FUNCTION_BLOCK LiftBootSync (* Basic Function Block Type *)
  (* Standard: 61499-2 *)
  (* Version 0.0, 11/25/2026, Schneider Electric, Sync Testing.Lift IRsp setpoint to resting sensor on boot *)
  PACKAGE Main;
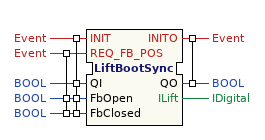
  EVENT_INPUT
    INIT WITH QI, FbOpen, FbClosed; (* Initialization Request *)
    REQ_FB_POS WITH FbOpen, FbClosed; (* Update Lift end-position feedback *)
  END_EVENT
  EVENT_OUTPUT
    INITO WITH QO; (* Initialization Confirm *)
  END_EVENT
  VAR_INPUT
    QI : BOOL := TRUE; (* Input event qualifier *)
    FbOpen : BOOL := FALSE; (* Lift raised end switch (1B1) *)
    FbClosed : BOOL := FALSE; (* Lift lowered end switch (1B2) *)
  END_VAR
  VAR_OUTPUT
    QO : BOOL; (* Output event qualifier *)
  END_VAR
  PLUGS
    ILift : IDigital; (* Remote setpoint adapter for Lift Valve2Op *)
  END_PLUGS
  VAR
    synced : BOOL := FALSE; (* Initial boot position synchronized to Lift IRsp *)
    prevTrack : BOOL := FALSE; (* Previous Track state from Lift IRsp *)
    targetSp : INT := 0; (* Tracked remote setpoint for Lift IRsp *)
    wantSend : BOOL := FALSE; (* Pending ILift.REQ event flag *)
  END_VAR
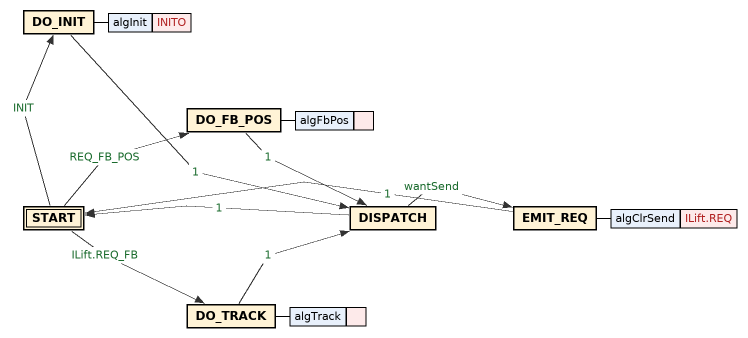
  EC_STATES
    START; (* Initial State *)
    DO_INIT : algInit -> INITO;
    DO_FB_POS : algFbPos;
    DO_TRACK : algTrack;
    DISPATCH;
    EMIT_REQ : algClrSend -> ILift.REQ;
  END_STATES
  EC_TRANSITIONS
    START TO DO_INIT := INIT;
    DO_INIT TO DISPATCH := 1;
    START TO DO_FB_POS := REQ_FB_POS;
    DO_FB_POS TO DISPATCH := 1;
    START TO DO_TRACK := ILift.REQ_FB;
    DO_TRACK TO DISPATCH := 1;
    DISPATCH TO EMIT_REQ := wantSend;
    EMIT_REQ TO START := 1;
    DISPATCH TO START := 1;
  END_TRANSITIONS
  ALGORITHM algInit IN ST: (* Initialize Lift boot sync state and match resting feedback if available *)
QO := QI;
synced := FALSE;
prevTrack := ILift.Track;
targetSp := 0;
wantSend := FALSE;
IF (NOT ILift.Track) AND (FbClosed OR FbOpen) THEN
	IF FbClosed AND NOT FbOpen THEN
		targetSp := 2;
		synced := TRUE;
		ILift.Value.value := targetSp;
		ILift.Value.quality := 16#0;
		wantSend := TRUE;
	ELSIF FbOpen AND NOT FbClosed THEN
		targetSp := 1;
		synced := TRUE;
		ILift.Value.value := targetSp;
		ILift.Value.quality := 16#0;
		wantSend := TRUE;
	END_IF;
END_IF;
  END_ALGORITHM
  ALGORITHM algFbPos IN ST: (* Sync initial IRsp setpoint to resting limit switch once on startup *)
IF (NOT synced) AND (NOT ILift.Track) AND (FbClosed OR FbOpen) THEN
	IF FbClosed AND NOT FbOpen THEN
		targetSp := 2;
		synced := TRUE;
		ILift.Value.value := targetSp;
		ILift.Value.quality := 16#0;
		wantSend := TRUE;
	ELSIF FbOpen AND NOT FbClosed THEN
		targetSp := 1;
		synced := TRUE;
		ILift.Value.value := targetSp;
		ILift.Value.quality := 16#0;
		wantSend := TRUE;
	END_IF;
END_IF;
  END_ALGORITHM
  ALGORITHM algTrack IN ST: (* Bumplessly track Operator/Program Local state and resync on return to Program Remote *)
IF ILift.Track THEN
	synced := TRUE;
	targetSp := ILift.State;
ELSIF prevTrack THEN
	synced := TRUE;
	ILift.Value.value := targetSp;
	ILift.Value.quality := 16#0;
	wantSend := TRUE;
ELSIF (NOT synced) AND (FbClosed OR FbOpen) THEN
	IF FbClosed AND NOT FbOpen THEN
		targetSp := 2;
		synced := TRUE;
		ILift.Value.value := targetSp;
		ILift.Value.quality := 16#0;
		wantSend := TRUE;
	ELSIF FbOpen AND NOT FbClosed THEN
		targetSp := 1;
		synced := TRUE;
		ILift.Value.value := targetSp;
		ILift.Value.quality := 16#0;
		wantSend := TRUE;
	END_IF;
END_IF;
prevTrack := ILift.Track;
  END_ALGORITHM
  ALGORITHM algClrSend IN ST: (* Clear pending ILift.REQ emit flag *)
wantSend := FALSE;
  END_ALGORITHM
END_FUNCTION_BLOCK
